{attribute 'GeneratedUsingTerminal: EK1100-0000-0018'}
{attribute addProperty BoxType "EK1100-0000-0018"}
{attribute addProperty Id "Term_280_EL1809EL1809_32157CFD20Term_281_EL1809EL1809_32157CFD20Term_282_EL1809EL1809_32157CFD20Term_283_EL1809EL1809_32157CFD20Term_284_EL1809EL1809_32157CFD20Term_312_EL1809EL1809_32157CFD20Term_320_EL1809EL1809_32157CFD20Term_321_EL1809EL1809_32157CFD20Term_322_EL1809EL1809_32157CFD20Term_323_EL1809EL1809_32157CFD20Term_324_EL1809EL1809_32157CFD20Term_325_EL1809EL1809_32157CFD20Term_326_EL1809EL1809_32157CFD20Term_327_EL1809EL1809_32157CFD20Term_328_EL1809EL1809_32157CFD20Term_329_EL1809EL1809_32157CFD20Term_331_EL1809EL1809_32157CFD20Term_332_EL1809EL1809_32157CFD20Term_333_EL1809EL1809_32157CFD20Term_334_EL1809EL1809_32157CFD20Term_335_EL1809EL1809_32157CFD20Term_336_EL1809EL1809_32157CFD20Term_337_EL1809EL1809_32157CFD20Term_338_EL1809EL1809_32157CFD20Term_339_EL1809EL1809_32157CFD20Term_340_EL1809EL1809_32157CFD20Term_341_EL1809EL1809_32157CFD20Term_342_EL1809EL1809_32157CFD20Term_343_EL1809EL1809_32157CFD20Term_344_EL1809EL1809_32157CFD20Term_345_EL1809EL1809_32157CFD20Term_346_EL1809EL1809_32157CFD20Term_347_EL1809EL1809_32157CFD20Term_348_EL1809EL1809_32157CFD20Term_360_EL1809EL1809_32157CFD20Term_361_EL1809EL1809_32157CFD20Term_362_EL1809EL1809_32157CFD20Term_363_EL1809EL1809_32157CFD20Term_364_EL1809EL1809_32157CFD20Term_365_EL1809EL1809_32157CFD20Term_366_EL1809EL1809_32157CFD20Term_367_EL1809EL1809_32157CFD20Term_368_EL1809EL1809_32157CFD20Term_370_EL1809EL1809_32157CFD20Term_371_EL1809EL1809_32157CFD20Term_372_EL1809EL1809_32157CFD20Term_373_EL1809EL1809_32157CFD20Term_374_EL1809EL1809_32157CFD20Term_375_EL1809EL1809_32157CFD20Term_376_EL1809EL1809_32157CFD20Term_377_EL1809EL1809_32157CFD20Term_378_EL1809EL1809_32157CFD20Term_380_EL1809EL1809_32157CFD20Term_381_EL1809EL1809_32157CFD20Term_382_EL1809EL1809_32157CFD20Term_383_EL1809EL1809_32157CFD20Term_384_EL1809EL1809_32157CFD20Term_385_EL1809EL1809_32157CFD20Term_386_EL1809EL1809_32157CFD20Term_387_EL1809EL1809_32157CFD20Term_388_EL1809EL1809_32157CFD20Term_389_EL1809EL1809_32157CFD20Term_390_EL1809EL1809_32157CFD20Term_391_EL1809EL1809_32157CFD20Term_392_EL1809EL1809_32157CFD20Term_393_EL1809EL1809_32157CFD20Term_394_EL1809EL1809_32157CFD20Term_395_EL1809EL1809_32157CFD20Term_396_EL1809EL1809_32157CFD20Term_397_EL1809EL1809_32157CFD20Term_398_EL1809EL1809_32157CFD20Term_399_EL1809EL1809_32157CFD20Term_400_EL1809EL1809_32157CFD20Term_401_EL1809EL1809_32157CFD20Term_402_EL1809EL1809_32157CFD20Term_403_EL1809EL1809_32157CFD20Term_404_EL1809EL1809_32157CFD20Term_405_EL1809EL1809_32157CFD20Term_406_EL1809EL1809_32157CFD20Term_407_EL1809EL1809_32157CFD20Term_408_EL1809EL1809_32157CFD20Term_409_EL1809EL1809_32157CFD20Term_410_EL1809EL1809_32157CFD20Term_414_EL1809EL1809_32157CFD20Term_415_EL1809EL1809_32157CFD20Term_416_EL1809EL1809_32157CFD20Term_417_EL1809EL1809_32157CFD20Term_418_EL1809EL1809_32157CFD20Term_419_EL1809EL1809_32157CFD20Term_420_EL1809EL1809_32157CFD20Term_421_EL1809EL1809_32157CFD20Term_422_EL1809EL1809_32157CFD20Term_423_EL1809EL1809_32157CFD20Term_424_EL1809EL1809_32157CFD20Term_425_EL1809EL1809_32157CFD20Term_426_EL1809EL1809_32157CFD20Term_427_EL1809EL1809_32157CFD20Term_428_EL1809EL1809_32157CFD20Term_429_EL1809EL1809_32157CFD20Term_448_EL1809EL1809_32157CFD20Term_495_EK1110EK1110_1FC0878B2"}
{attribute addProperty CRC "3984417394"}
{attribute addProperty Size "2002"}
{attribute addProperty Name "Term 279 (EK1100)"}
TYPE Term_279_EK1100_ED7D6272 EXTENDS EK1100_1FC0878B :
STRUCT
	{attribute addProperty Name "Term 280 (EL1809)"}
	{attribute addProperty PreviousPort "Term 279 (EK1100) : B"}
	{attribute addProperty SyncUnit "default"}
	Term_280_EL1809 : EL1809_32157CFD;
	{attribute addProperty Name "Term 281 (EL1809)"}
	{attribute addProperty PreviousPort "Term 280 (EL1809) : B"}
	{attribute addProperty SyncUnit "default"}
	Term_281_EL1809 : EL1809_32157CFD;
	{attribute addProperty Name "Term 282 (EL1809)"}
	{attribute addProperty PreviousPort "Term 281 (EL1809) : B"}
	{attribute addProperty SyncUnit "default"}
	Term_282_EL1809 : EL1809_32157CFD;
	{attribute addProperty Name "Term 283 (EL1809)"}
	{attribute addProperty PreviousPort "Term 282 (EL1809) : B"}
	{attribute addProperty SyncUnit "default"}
	Term_283_EL1809 : EL1809_32157CFD;
	{attribute addProperty Name "Term 284 (EL1809)"}
	{attribute addProperty PreviousPort "Term 283 (EL1809) : B"}
	{attribute addProperty SyncUnit "default"}
	Term_284_EL1809 : EL1809_32157CFD;
	{attribute addProperty Name "Term 312 (EL1809)"}
	{attribute addProperty PreviousPort "Term 284 (EL1809) : B"}
	{attribute addProperty SyncUnit "default"}
	Term_312_EL1809 : EL1809_32157CFD;
	{attribute addProperty Name "Term 320 (EL1809)"}
	{attribute addProperty PreviousPort "Term 312 (EL1809) : B"}
	{attribute addProperty SyncUnit "default"}
	Term_320_EL1809 : EL1809_32157CFD;
	{attribute addProperty Name "Term 321 (EL1809)"}
	{attribute addProperty PreviousPort "Term 320 (EL1809) : B"}
	{attribute addProperty SyncUnit "default"}
	Term_321_EL1809 : EL1809_32157CFD;
	{attribute addProperty Name "Term 322 (EL1809)"}
	{attribute addProperty PreviousPort "Term 321 (EL1809) : B"}
	{attribute addProperty SyncUnit "default"}
	Term_322_EL1809 : EL1809_32157CFD;
	{attribute addProperty Name "Term 323 (EL1809)"}
	{attribute addProperty PreviousPort "Term 322 (EL1809) : B"}
	{attribute addProperty SyncUnit "default"}
	Term_323_EL1809 : EL1809_32157CFD;
	{attribute addProperty Name "Term 324 (EL1809)"}
	{attribute addProperty PreviousPort "Term 323 (EL1809) : B"}
	{attribute addProperty SyncUnit "default"}
	Term_324_EL1809 : EL1809_32157CFD;
	{attribute addProperty Name "Term 325 (EL1809)"}
	{attribute addProperty PreviousPort "Term 324 (EL1809) : B"}
	{attribute addProperty SyncUnit "default"}
	Term_325_EL1809 : EL1809_32157CFD;
	{attribute addProperty Name "Term 326 (EL1809)"}
	{attribute addProperty PreviousPort "Term 325 (EL1809) : B"}
	{attribute addProperty SyncUnit "default"}
	Term_326_EL1809 : EL1809_32157CFD;
	{attribute addProperty Name "Term 327 (EL1809)"}
	{attribute addProperty PreviousPort "Term 326 (EL1809) : B"}
	{attribute addProperty SyncUnit "default"}
	Term_327_EL1809 : EL1809_32157CFD;
	{attribute addProperty Name "Term 328 (EL1809)"}
	{attribute addProperty PreviousPort "Term 327 (EL1809) : B"}
	{attribute addProperty SyncUnit "default"}
	Term_328_EL1809 : EL1809_32157CFD;
	{attribute addProperty Name "Term 329 (EL1809)"}
	{attribute addProperty PreviousPort "Term 328 (EL1809) : B"}
	{attribute addProperty SyncUnit "default"}
	Term_329_EL1809 : EL1809_32157CFD;
	{attribute addProperty Name "Term 331 (EL1809)"}
	{attribute addProperty PreviousPort "Term 329 (EL1809) : B"}
	{attribute addProperty SyncUnit "default"}
	Term_331_EL1809 : EL1809_32157CFD;
	{attribute addProperty Name "Term 332 (EL1809)"}
	{attribute addProperty PreviousPort "Term 331 (EL1809) : B"}
	{attribute addProperty SyncUnit "default"}
	Term_332_EL1809 : EL1809_32157CFD;
	{attribute addProperty Name "Term 333 (EL1809)"}
	{attribute addProperty PreviousPort "Term 332 (EL1809) : B"}
	{attribute addProperty SyncUnit "default"}
	Term_333_EL1809 : EL1809_32157CFD;
	{attribute addProperty Name "Term 334 (EL1809)"}
	{attribute addProperty PreviousPort "Term 333 (EL1809) : B"}
	{attribute addProperty SyncUnit "default"}
	Term_334_EL1809 : EL1809_32157CFD;
	{attribute addProperty Name "Term 335 (EL1809)"}
	{attribute addProperty PreviousPort "Term 334 (EL1809) : B"}
	{attribute addProperty SyncUnit "default"}
	Term_335_EL1809 : EL1809_32157CFD;
	{attribute addProperty Name "Term 336 (EL1809)"}
	{attribute addProperty PreviousPort "Term 335 (EL1809) : B"}
	{attribute addProperty SyncUnit "default"}
	Term_336_EL1809 : EL1809_32157CFD;
	{attribute addProperty Name "Term 337 (EL1809)"}
	{attribute addProperty PreviousPort "Term 336 (EL1809) : B"}
	{attribute addProperty SyncUnit "default"}
	Term_337_EL1809 : EL1809_32157CFD;
	{attribute addProperty Name "Term 338 (EL1809)"}
	{attribute addProperty PreviousPort "Term 337 (EL1809) : B"}
	{attribute addProperty SyncUnit "default"}
	Term_338_EL1809 : EL1809_32157CFD;
	{attribute addProperty Name "Term 339 (EL1809)"}
	{attribute addProperty PreviousPort "Term 338 (EL1809) : B"}
	{attribute addProperty SyncUnit "default"}
	Term_339_EL1809 : EL1809_32157CFD;
	{attribute addProperty Name "Term 340 (EL1809)"}
	{attribute addProperty PreviousPort "Term 339 (EL1809) : B"}
	{attribute addProperty SyncUnit "default"}
	Term_340_EL1809 : EL1809_32157CFD;
	{attribute addProperty Name "Term 341 (EL1809)"}
	{attribute addProperty PreviousPort "Term 340 (EL1809) : B"}
	{attribute addProperty SyncUnit "default"}
	Term_341_EL1809 : EL1809_32157CFD;
	{attribute addProperty Name "Term 342 (EL1809)"}
	{attribute addProperty PreviousPort "Term 341 (EL1809) : B"}
	{attribute addProperty SyncUnit "default"}
	Term_342_EL1809 : EL1809_32157CFD;
	{attribute addProperty Name "Term 343 (EL1809)"}
	{attribute addProperty PreviousPort "Term 342 (EL1809) : B"}
	{attribute addProperty SyncUnit "default"}
	Term_343_EL1809 : EL1809_32157CFD;
	{attribute addProperty Name "Term 344 (EL1809)"}
	{attribute addProperty PreviousPort "Term 343 (EL1809) : B"}
	{attribute addProperty SyncUnit "default"}
	Term_344_EL1809 : EL1809_32157CFD;
	{attribute addProperty Name "Term 345 (EL1809)"}
	{attribute addProperty PreviousPort "Term 344 (EL1809) : B"}
	{attribute addProperty SyncUnit "default"}
	Term_345_EL1809 : EL1809_32157CFD;
	{attribute addProperty Name "Term 346 (EL1809)"}
	{attribute addProperty PreviousPort "Term 345 (EL1809) : B"}
	{attribute addProperty SyncUnit "default"}
	Term_346_EL1809 : EL1809_32157CFD;
	{attribute addProperty Name "Term 347 (EL1809)"}
	{attribute addProperty PreviousPort "Term 346 (EL1809) : B"}
	{attribute addProperty SyncUnit "default"}
	Term_347_EL1809 : EL1809_32157CFD;
	{attribute addProperty Name "Term 348 (EL1809)"}
	{attribute addProperty PreviousPort "Term 347 (EL1809) : B"}
	{attribute addProperty SyncUnit "default"}
	Term_348_EL1809 : EL1809_32157CFD;
	{attribute addProperty Name "Term 360 (EL1809)"}
	{attribute addProperty PreviousPort "Term 348 (EL1809) : B"}
	{attribute addProperty SyncUnit "default"}
	Term_360_EL1809 : EL1809_32157CFD;
	{attribute addProperty Name "Term 361 (EL1809)"}
	{attribute addProperty PreviousPort "Term 360 (EL1809) : B"}
	{attribute addProperty SyncUnit "default"}
	Term_361_EL1809 : EL1809_32157CFD;
	{attribute addProperty Name "Term 362 (EL1809)"}
	{attribute addProperty PreviousPort "Term 361 (EL1809) : B"}
	{attribute addProperty SyncUnit "default"}
	Term_362_EL1809 : EL1809_32157CFD;
	{attribute addProperty Name "Term 363 (EL1809)"}
	{attribute addProperty PreviousPort "Term 362 (EL1809) : B"}
	{attribute addProperty SyncUnit "default"}
	Term_363_EL1809 : EL1809_32157CFD;
	{attribute addProperty Name "Term 364 (EL1809)"}
	{attribute addProperty PreviousPort "Term 363 (EL1809) : B"}
	{attribute addProperty SyncUnit "default"}
	Term_364_EL1809 : EL1809_32157CFD;
	{attribute addProperty Name "Term 365 (EL1809)"}
	{attribute addProperty PreviousPort "Term 364 (EL1809) : B"}
	{attribute addProperty SyncUnit "default"}
	Term_365_EL1809 : EL1809_32157CFD;
	{attribute addProperty Name "Term 366 (EL1809)"}
	{attribute addProperty PreviousPort "Term 365 (EL1809) : B"}
	{attribute addProperty SyncUnit "default"}
	Term_366_EL1809 : EL1809_32157CFD;
	{attribute addProperty Name "Term 367 (EL1809)"}
	{attribute addProperty PreviousPort "Term 366 (EL1809) : B"}
	{attribute addProperty SyncUnit "default"}
	Term_367_EL1809 : EL1809_32157CFD;
	{attribute addProperty Name "Term 368 (EL1809)"}
	{attribute addProperty PreviousPort "Term 367 (EL1809) : B"}
	{attribute addProperty SyncUnit "default"}
	Term_368_EL1809 : EL1809_32157CFD;
	{attribute addProperty Name "Term 370 (EL1809)"}
	{attribute addProperty PreviousPort "Term 368 (EL1809) : B"}
	{attribute addProperty SyncUnit "default"}
	Term_370_EL1809 : EL1809_32157CFD;
	{attribute addProperty Name "Term 371 (EL1809)"}
	{attribute addProperty PreviousPort "Term 370 (EL1809) : B"}
	{attribute addProperty SyncUnit "default"}
	Term_371_EL1809 : EL1809_32157CFD;
	{attribute addProperty Name "Term 372 (EL1809)"}
	{attribute addProperty PreviousPort "Term 371 (EL1809) : B"}
	{attribute addProperty SyncUnit "default"}
	Term_372_EL1809 : EL1809_32157CFD;
	{attribute addProperty Name "Term 373 (EL1809)"}
	{attribute addProperty PreviousPort "Term 372 (EL1809) : B"}
	{attribute addProperty SyncUnit "default"}
	Term_373_EL1809 : EL1809_32157CFD;
	{attribute addProperty Name "Term 374 (EL1809)"}
	{attribute addProperty PreviousPort "Term 373 (EL1809) : B"}
	{attribute addProperty SyncUnit "default"}
	Term_374_EL1809 : EL1809_32157CFD;
	{attribute addProperty Name "Term 375 (EL1809)"}
	{attribute addProperty PreviousPort "Term 374 (EL1809) : B"}
	{attribute addProperty SyncUnit "default"}
	Term_375_EL1809 : EL1809_32157CFD;
	{attribute addProperty Name "Term 376 (EL1809)"}
	{attribute addProperty PreviousPort "Term 375 (EL1809) : B"}
	{attribute addProperty SyncUnit "default"}
	Term_376_EL1809 : EL1809_32157CFD;
	{attribute addProperty Name "Term 377 (EL1809)"}
	{attribute addProperty PreviousPort "Term 376 (EL1809) : B"}
	{attribute addProperty SyncUnit "default"}
	Term_377_EL1809 : EL1809_32157CFD;
	{attribute addProperty Name "Term 378 (EL1809)"}
	{attribute addProperty PreviousPort "Term 377 (EL1809) : B"}
	{attribute addProperty SyncUnit "default"}
	Term_378_EL1809 : EL1809_32157CFD;
	{attribute addProperty Name "Term 380 (EL1809)"}
	{attribute addProperty PreviousPort "Term 378 (EL1809) : B"}
	{attribute addProperty SyncUnit "default"}
	Term_380_EL1809 : EL1809_32157CFD;
	{attribute addProperty Name "Term 381 (EL1809)"}
	{attribute addProperty PreviousPort "Term 380 (EL1809) : B"}
	{attribute addProperty SyncUnit "default"}
	Term_381_EL1809 : EL1809_32157CFD;
	{attribute addProperty Name "Term 382 (EL1809)"}
	{attribute addProperty PreviousPort "Term 381 (EL1809) : B"}
	{attribute addProperty SyncUnit "default"}
	Term_382_EL1809 : EL1809_32157CFD;
	{attribute addProperty Name "Term 383 (EL1809)"}
	{attribute addProperty PreviousPort "Term 382 (EL1809) : B"}
	{attribute addProperty SyncUnit "default"}
	Term_383_EL1809 : EL1809_32157CFD;
	{attribute addProperty Name "Term 384 (EL1809)"}
	{attribute addProperty PreviousPort "Term 383 (EL1809) : B"}
	{attribute addProperty SyncUnit "default"}
	Term_384_EL1809 : EL1809_32157CFD;
	{attribute addProperty Name "Term 385 (EL1809)"}
	{attribute addProperty PreviousPort "Term 384 (EL1809) : B"}
	{attribute addProperty SyncUnit "default"}
	Term_385_EL1809 : EL1809_32157CFD;
	{attribute addProperty Name "Term 386 (EL1809)"}
	{attribute addProperty PreviousPort "Term 385 (EL1809) : B"}
	{attribute addProperty SyncUnit "default"}
	Term_386_EL1809 : EL1809_32157CFD;
	{attribute addProperty Name "Term 387 (EL1809)"}
	{attribute addProperty PreviousPort "Term 386 (EL1809) : B"}
	{attribute addProperty SyncUnit "default"}
	Term_387_EL1809 : EL1809_32157CFD;
	{attribute addProperty Name "Term 388 (EL1809)"}
	{attribute addProperty PreviousPort "Term 387 (EL1809) : B"}
	{attribute addProperty SyncUnit "default"}
	Term_388_EL1809 : EL1809_32157CFD;
	{attribute addProperty Name "Term 389 (EL1809)"}
	{attribute addProperty PreviousPort "Term 388 (EL1809) : B"}
	{attribute addProperty SyncUnit "default"}
	Term_389_EL1809 : EL1809_32157CFD;
	{attribute addProperty Name "Term 390 (EL1809)"}
	{attribute addProperty PreviousPort "Term 389 (EL1809) : B"}
	{attribute addProperty SyncUnit "default"}
	Term_390_EL1809 : EL1809_32157CFD;
	{attribute addProperty Name "Term 391 (EL1809)"}
	{attribute addProperty PreviousPort "Term 390 (EL1809) : B"}
	{attribute addProperty SyncUnit "default"}
	Term_391_EL1809 : EL1809_32157CFD;
	{attribute addProperty Name "Term 392 (EL1809)"}
	{attribute addProperty PreviousPort "Term 391 (EL1809) : B"}
	{attribute addProperty SyncUnit "default"}
	Term_392_EL1809 : EL1809_32157CFD;
	{attribute addProperty Name "Term 393 (EL1809)"}
	{attribute addProperty PreviousPort "Term 392 (EL1809) : B"}
	{attribute addProperty SyncUnit "default"}
	Term_393_EL1809 : EL1809_32157CFD;
	{attribute addProperty Name "Term 394 (EL1809)"}
	{attribute addProperty PreviousPort "Term 393 (EL1809) : B"}
	{attribute addProperty SyncUnit "default"}
	Term_394_EL1809 : EL1809_32157CFD;
	{attribute addProperty Name "Term 395 (EL1809)"}
	{attribute addProperty PreviousPort "Term 394 (EL1809) : B"}
	{attribute addProperty SyncUnit "default"}
	Term_395_EL1809 : EL1809_32157CFD;
	{attribute addProperty Name "Term 396 (EL1809)"}
	{attribute addProperty PreviousPort "Term 395 (EL1809) : B"}
	{attribute addProperty SyncUnit "default"}
	Term_396_EL1809 : EL1809_32157CFD;
	{attribute addProperty Name "Term 397 (EL1809)"}
	{attribute addProperty PreviousPort "Term 396 (EL1809) : B"}
	{attribute addProperty SyncUnit "default"}
	Term_397_EL1809 : EL1809_32157CFD;
	{attribute addProperty Name "Term 398 (EL1809)"}
	{attribute addProperty PreviousPort "Term 397 (EL1809) : B"}
	{attribute addProperty SyncUnit "default"}
	Term_398_EL1809 : EL1809_32157CFD;
	{attribute addProperty Name "Term 399 (EL1809)"}
	{attribute addProperty PreviousPort "Term 398 (EL1809) : B"}
	{attribute addProperty SyncUnit "default"}
	Term_399_EL1809 : EL1809_32157CFD;
	{attribute addProperty Name "Term 400 (EL1809)"}
	{attribute addProperty PreviousPort "Term 399 (EL1809) : B"}
	{attribute addProperty SyncUnit "default"}
	Term_400_EL1809 : EL1809_32157CFD;
	{attribute addProperty Name "Term 401 (EL1809)"}
	{attribute addProperty PreviousPort "Term 400 (EL1809) : B"}
	{attribute addProperty SyncUnit "default"}
	Term_401_EL1809 : EL1809_32157CFD;
	{attribute addProperty Name "Term 402 (EL1809)"}
	{attribute addProperty PreviousPort "Term 401 (EL1809) : B"}
	{attribute addProperty SyncUnit "default"}
	Term_402_EL1809 : EL1809_32157CFD;
	{attribute addProperty Name "Term 403 (EL1809)"}
	{attribute addProperty PreviousPort "Term 402 (EL1809) : B"}
	{attribute addProperty SyncUnit "default"}
	Term_403_EL1809 : EL1809_32157CFD;
	{attribute addProperty Name "Term 404 (EL1809)"}
	{attribute addProperty PreviousPort "Term 403 (EL1809) : B"}
	{attribute addProperty SyncUnit "default"}
	Term_404_EL1809 : EL1809_32157CFD;
	{attribute addProperty Name "Term 405 (EL1809)"}
	{attribute addProperty PreviousPort "Term 404 (EL1809) : B"}
	{attribute addProperty SyncUnit "default"}
	Term_405_EL1809 : EL1809_32157CFD;
	{attribute addProperty Name "Term 406 (EL1809)"}
	{attribute addProperty PreviousPort "Term 405 (EL1809) : B"}
	{attribute addProperty SyncUnit "default"}
	Term_406_EL1809 : EL1809_32157CFD;
	{attribute addProperty Name "Term 407 (EL1809)"}
	{attribute addProperty PreviousPort "Term 406 (EL1809) : B"}
	{attribute addProperty SyncUnit "default"}
	Term_407_EL1809 : EL1809_32157CFD;
	{attribute addProperty Name "Term 408 (EL1809)"}
	{attribute addProperty PreviousPort "Term 407 (EL1809) : B"}
	{attribute addProperty SyncUnit "default"}
	Term_408_EL1809 : EL1809_32157CFD;
	{attribute addProperty Name "Term 409 (EL1809)"}
	{attribute addProperty PreviousPort "Term 408 (EL1809) : B"}
	{attribute addProperty SyncUnit "default"}
	Term_409_EL1809 : EL1809_32157CFD;
	{attribute addProperty Name "Term 410 (EL1809)"}
	{attribute addProperty PreviousPort "Term 409 (EL1809) : B"}
	{attribute addProperty SyncUnit "default"}
	Term_410_EL1809 : EL1809_32157CFD;
	{attribute addProperty Name "Term 414 (EL1809)"}
	{attribute addProperty PreviousPort "Term 410 (EL1809) : B"}
	{attribute addProperty SyncUnit "default"}
	Term_414_EL1809 : EL1809_32157CFD;
	{attribute addProperty Name "Term 415 (EL1809)"}
	{attribute addProperty PreviousPort "Term 414 (EL1809) : B"}
	{attribute addProperty SyncUnit "default"}
	Term_415_EL1809 : EL1809_32157CFD;
	{attribute addProperty Name "Term 416 (EL1809)"}
	{attribute addProperty PreviousPort "Term 415 (EL1809) : B"}
	{attribute addProperty SyncUnit "default"}
	Term_416_EL1809 : EL1809_32157CFD;
	{attribute addProperty Name "Term 417 (EL1809)"}
	{attribute addProperty PreviousPort "Term 416 (EL1809) : B"}
	{attribute addProperty SyncUnit "default"}
	Term_417_EL1809 : EL1809_32157CFD;
	{attribute addProperty Name "Term 418 (EL1809)"}
	{attribute addProperty PreviousPort "Term 417 (EL1809) : B"}
	{attribute addProperty SyncUnit "default"}
	Term_418_EL1809 : EL1809_32157CFD;
	{attribute addProperty Name "Term 419 (EL1809)"}
	{attribute addProperty PreviousPort "Term 418 (EL1809) : B"}
	{attribute addProperty SyncUnit "default"}
	Term_419_EL1809 : EL1809_32157CFD;
	{attribute addProperty Name "Term 420 (EL1809)"}
	{attribute addProperty PreviousPort "Term 419 (EL1809) : B"}
	{attribute addProperty SyncUnit "default"}
	Term_420_EL1809 : EL1809_32157CFD;
	{attribute addProperty Name "Term 421 (EL1809)"}
	{attribute addProperty PreviousPort "Term 420 (EL1809) : B"}
	{attribute addProperty SyncUnit "default"}
	Term_421_EL1809 : EL1809_32157CFD;
	{attribute addProperty Name "Term 422 (EL1809)"}
	{attribute addProperty PreviousPort "Term 421 (EL1809) : B"}
	{attribute addProperty SyncUnit "default"}
	Term_422_EL1809 : EL1809_32157CFD;
	{attribute addProperty Name "Term 423 (EL1809)"}
	{attribute addProperty PreviousPort "Term 422 (EL1809) : B"}
	{attribute addProperty SyncUnit "default"}
	Term_423_EL1809 : EL1809_32157CFD;
	{attribute addProperty Name "Term 424 (EL1809)"}
	{attribute addProperty PreviousPort "Term 423 (EL1809) : B"}
	{attribute addProperty SyncUnit "default"}
	Term_424_EL1809 : EL1809_32157CFD;
	{attribute addProperty Name "Term 425 (EL1809)"}
	{attribute addProperty PreviousPort "Term 424 (EL1809) : B"}
	{attribute addProperty SyncUnit "default"}
	Term_425_EL1809 : EL1809_32157CFD;
	{attribute addProperty Name "Term 426 (EL1809)"}
	{attribute addProperty PreviousPort "Term 425 (EL1809) : B"}
	{attribute addProperty SyncUnit "default"}
	Term_426_EL1809 : EL1809_32157CFD;
	{attribute addProperty Name "Term 427 (EL1809)"}
	{attribute addProperty PreviousPort "Term 426 (EL1809) : B"}
	{attribute addProperty SyncUnit "default"}
	Term_427_EL1809 : EL1809_32157CFD;
	{attribute addProperty Name "Term 428 (EL1809)"}
	{attribute addProperty PreviousPort "Term 427 (EL1809) : B"}
	{attribute addProperty SyncUnit "default"}
	Term_428_EL1809 : EL1809_32157CFD;
	{attribute addProperty Name "Term 429 (EL1809)"}
	{attribute addProperty PreviousPort "Term 428 (EL1809) : B"}
	{attribute addProperty SyncUnit "default"}
	Term_429_EL1809 : EL1809_32157CFD;
	{attribute addProperty Name "Term 448 (EL1809)"}
	{attribute addProperty PreviousPort "Term 429 (EL1809) : B"}
	{attribute addProperty SyncUnit "default"}
	Term_448_EL1809 : EL1809_32157CFD;
	{attribute addProperty Name "Term 495 (EK1110)"}
	{attribute addProperty PreviousPort "Term 448 (EL1809) : B"}
	{attribute addProperty SyncUnit "default"}
	Term_495_EK1110 : EK1110_1FC0878B;
END_STRUCT
END_TYPE

(* stored: Version 1.2.0.0, ProductVersion 3.1.4024.11
   DUT Term_279_EK1100_ED7D6272: Id {1570f905-b890-0d43-0174-4a551da94df0} *)
